// SIMATIC S7-200 SMART project (STEP 7-Micro/WIN SMART), CPU ST40

SYMBOL_TABLE ACTUATOR MEMORY
X_EXTEND         M2.0     // X EXTEND
X_RETRACT        M2.1     // X RETRACT
Y_EXTEND         M2.2     // Y EXTEND
Y_RETRACT        M2.3     // Y RETRACT
Z_EXTEND         M2.4     // Z EXTEND
Z_RETRACT        M2.5     // Z RETRACT
GRIPPER          M2.6     // GRIPPER
END_SYMBOL_TABLE

SYMBOL_TABLE System Symbols
ON_STATE         M0.0     // ON STATE
END_SYMBOL_TABLE

SYMBOL_TABLE STEPS MEMORY
STEP_1_START     M1.0     // STEP 1 ONLINE
END_SYMBOL_TABLE

SYMBOL_TABLE MOVEMENT MEMORY
X_MOVEMENT       M3.0     // X_MOVEMENT
Y_MOVEMENT       M3.1     // Y_MOVEMENT
Z_MOVEMENT       M3.2     // Z_MOVEMENT
GRIPPER_MOVEMENT M3.3     // GRIPPER_MOVEMENT
END_SYMBOL_TABLE

ORGANIZATION_BLOCK MAIN:OB1
TITLE=Program Comments
BEGIN
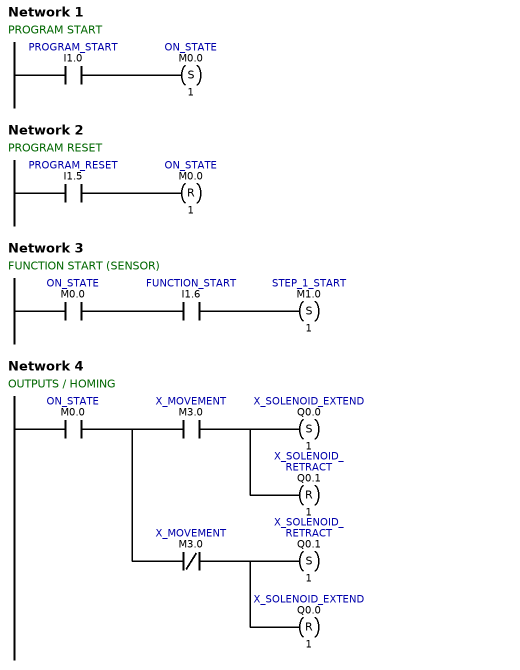
Network 1
// PROGRAM START
LD     PROGRAM_START:I1.0
S      ON_STATE:M0.0, 1
Network 2
// PROGRAM RESET
LD     PROGRAM_RESET:I1.5
R      ON_STATE:M0.0, 1
Network 3
// FUNCTION START (SENSOR)
LD     ON_STATE:M0.0
A      FUNCTION_START:I1.6
S      STEP_1_START:M1.0, 1
Network 4
// OUTPUTS / HOMING
LD     ON_STATE:M0.0
LPS
A      X_MOVEMENT:M3.0
S      X_SOLENOID_EXTEND:Q0.0, 1
R      X_SOLENOID_RETRACT:Q0.1, 1
LPP
AN     X_MOVEMENT:M3.0
S      X_SOLENOID_RETRACT:Q0.1, 1
R      X_SOLENOID_EXTEND:Q0.0, 1
Network 5
// MEMORY MOVEMENT
// 
END_ORGANIZATION_BLOCK
